(*
SPDX-FileCopyrightText: © 2026 Oleksandr Tiutyk <trofimich@gmail.com>
SPDX-License-Identifier: MIT
License: https://opensource.org/license/mit
*)

(*!
<summary>Identifies an optional domain-specific deserialization context queried during deserialization.</summary>
<description>
Marker interface without members. Passed to IConfigurationSerializable.Deserialize for the duration of a
single synchronous call to supply domain-specific reconstruction services (such as workflow element loaders or
dependency resolvers) queried via __QUERYINTERFACE.
The context is borrowed and must not be retained or stored by the deserialized object across execution cycles.
A null context (context = 0) is valid when no external services are available. Objects requiring specific
context capabilities must validate the context explicitly and raise a configuration exception when absent or
incompatible.
</description>
*)
INTERFACE IConfigurationDeserializationContext EXTENDS IObject

END_INTERFACE

(* stored: Version 1.1.0.1
   Itf IConfigurationDeserializationContext: Id {f261b8da-6be1-41ed-bfe6-3a3ff28eb591} *)
